Fanuc KAREL source: ka00056.KL

-- PROVISIONAL review KL for V1013-1; original PC SHA256 f5c90b6702f43ddaf0e01a470d18fb833bafcc281b8aba1152de6eae93bd0056
-- Incomplete behavior may be omitted. Consult companion uncertainty JSON. Do not deploy.
PROGRAM KA00056
%NOLOCKGROUP
-- UNRESOLVED_DECL SRC type=000101
-- UNRESOLVED_DECL DST type=000199
BEGIN
  -- UNRESOLVED_PC offsets 5-25; opcodes 49,7E,4A
  -- UNRESOLVED_PC offsets 30-34; opcodes 7F
END KA00056
